(* IEC 61131-3 sources: Gen-AI/docs/member2_validation/codesys_release_v1.1/C05_dead_code, 1 file *)

(* ---- source.st ---- *)
FUNCTION_BLOCK FB_AgentProbeDeadCode
VAR_OUTPUT
 y : BOOL;
END_VAR
IF FALSE THEN
 y := TRUE;
ELSE
 y := FALSE;
END_IF;
END_FUNCTION_BLOCK
